(* IEC 61131-3 sources: Test-Git_ESME26/TestProgettoESME_26.fbsproj/PacDriveLib_Motion_Migration_Example.device.xml.v3^/Plc Logic.plclogic.xml.v3^/Application.application.xml.v3^/Test_MultiCam, 1 file *)

(* ---- GVL_Encoder.gvl ---- *)
VAR_GLOBAL
	Logical_Encoder				: MOIN.FB_LogicalEncoder;
	Logical_Encoder_YOffset		: MOIN.FB_LogicalEncoder;
END_VAR
